// TIA Portal V20 export
// export: Created 2026-10-19T18:45:37.2686399Z, ExportSetting None, DisplayName Totally Integrated Automation Portal, DisplayVersion V20 Update 6, DisplayName TIA Portal Openness, DisplayVersion V20 Update 6, DisplayName TIA Portal Version Control Interface, DisplayVersion V20 Update 6, DisplayName SINAMICS Startdrive Advanced, DisplayVersion V20 SP1, DisplayName SINAMICS Startdrive G130, G150, S120, S150, SINAMICS MV, G220, S200, S210, DisplayVersion V20 SP1, DisplayName SINAMICS Startdrive G110M, G120, G120C, G120D, G120P, G115D, DisplayVersion V20 SP1, DisplayName STEP 7 Professional, DisplayVersion V20 Update 6, DisplayName STEP 7 Safety, DisplayVersion V20 Update 2, DisplayName WinCC Basic/Comfort/Advanced, DisplayVersion V20 Update 6, DisplayName WinCC Unified, DisplayVersion V20 Update 6
VAR_GLOBAL   // PLC tag table "IO_Remote_Panel_2"
   "KEY REMOTE/LOCAL L5 - CH1(2)" AT %I470.5 : Bool;
   "KEY REMOTE/LOCAL L2 - CH1(2)" AT %I461.7 : Bool;
   "VTD2 UPPER ULTIMATE CREEP" AT %I286.1 : Bool;
   "SAFETY_GATE_3_CH1(2)" AT %I461.2 : Bool;
   "STACK LIGHTS GREEN(2)" AT %Q174.3 : Bool;
   "C2112 VTD CIRCUIT BREAKER" AT %I285.0 : Bool;
   "STO VTD - CH1(2)" AT %Q446.2 : Bool;
   "STACK LIGHTS RED(2)" AT %Q174.1 : Bool;
   "LIGHT GUARDS 2 - CH2(2)" AT %I453.2 : Bool;
   "VTU HOIST BRAKE SAFETY ENABLE EDM FEEDBACK(2)" AT %I452.0 : Bool;
   "Chain Slack 3 - CH1(2)" AT %I356.6 : Bool;
   "KEY REMOTE/LOCAL L3 - CH1(2)" AT %I470.1 : Bool;
   "KEY REMOTE/LOCAL L6 - CH1(2)" AT %I470.7 : Bool;
   "BRAKE SUPPLY SAFETY CONTACTOR 1(2)" AT %Q446.0 : Bool;
   "KEY REMOTE/LOCAL L1 - CH2(2)" AT %I462.5 : Bool;
   "E-STOP L1 - CH2(2)" AT %I462.4 : Bool;
   "E-STOP L1 - CH1(2)" AT %I461.4 : Bool;
   "VTD2 PUSH TO EXIT VTD ZONE" AT %I286.6 : Bool;
   "E-STOP (CABINET) - CH1(2)" AT %I356.0 : Bool;
   "E-STOP L6 - CH2(2)" AT %I471.6 : Bool;
   "C2109, C2110, C2111 CVTD CIRCUIT BREAKER" AT %I285.3 : Bool;
   "E-STOP L2 - CH2(2)" AT %I462.6 : Bool;
   "SAFETY_GATE_1_CH2(2)" AT %I462.0 : Bool;
   "CABINET COOLING FAN CIRCUIT BREAKER FEEDBACK(2)" AT %I285.4 : Bool;
   "KEY REMOTE/LOCAL L6 - CH2(2)" AT %I471.7 : Bool;
   "STO VTD - CH2(2)" AT %Q446.3 : Bool;
   "KEY REMOTE/LOCAL L1 - CH1(2)" AT %I461.5 : Bool;
   "SAFETY_GATE_1_CH1(2)" AT %I461.0 : Bool;
   "KEY REMOTE/LOCAL L3 - CH2(2)" AT %I471.1 : Bool;
   "VTD2 UPPER ULTIMATE SLOWDOWN" AT %I286.0 : Bool;
   "VTD2 LOWER ULTIMATE SLOWDOWN" AT %I286.4 : Bool;
   "KEY REMOTE/LOCAL L4 - CH2(2)" AT %I471.3 : Bool;
   "E-STOP L6 - CH1(2)" AT %I470.6 : Bool;
   "KEY REMOTE/LOCAL L4 - CH1(2)" AT %I470.3 : Bool;
   "E-STOP L5 - CH1(2)" AT %I470.4 : Bool;
   "E-STOP L3 - CH2(2)" AT %I471.0 : Bool;
   "KEY REMOTE/LOCAL L5 - CH2(2)" AT %I471.5 : Bool;
   "BRAKE SUPPLY SAFETY CONTACTOR 2(2)" AT %Q446.1 : Bool;
   "SAFETY_GATE_4_CH1(2)" AT %I461.3 : Bool;
   "Chain Slack 3 - CH2(2)" AT %I357.6 : Bool;
   "STACK LIGHTS ORANGE(2)" AT %Q174.2 : Bool;
   "Chain Slack 2 - CH2(2)" AT %I357.5 : Bool;
   "C2105, C2106, C2107, C2108 CIRCUIT BREAKER" AT %I285.2 : Bool;
   "LIGHT GUARD 2 - CH1(2)" AT %I452.2 : Bool;
   "Chain Slack 2 - CH1(2)" AT %I356.5 : Bool;
   "KEY REMOTE/LOCAL L2 - CH2(2)" AT %I462.7 : Bool;
   "VTD2 PUSH TO ENTER VTD ZONE" AT %I286.5 : Bool;
   "CABINET 24V PSU CIRCUIT BREAKER FEEDBACK(2)" AT %I285.5 : Bool;
   "CABINET 24V PSU CIRCUIT BREAKER FEEDBACK_1(2)" AT %I285.6 : Bool;
   "Chain Slack 1 - CH1(2)" AT %I356.4 : Bool;
   "SAFETY_GATE_3_CH2(2)" AT %I462.2 : Bool;
   "RESET (CABINET)(2)" AT %I356.1 : Bool;
   "E-STOP L3 - CH1(2)" AT %I470.0 : Bool;
   "RESET LAMP(2)" AT %Q174.0 : Bool;   // TESTED
   "SAFETY_GATE_2_CH1(2)" AT %I461.1 : Bool;
   "E-STOP L5 - CH2(2)" AT %I471.4 : Bool;
   "VTD2 UPPER LIMIT" AT %I286.3 : Bool;
   "LIGHT GUARDS 1 - CH2(2)" AT %I453.1 : Bool;
   "Chain Slack 1 - CH2(2)" AT %I357.4 : Bool;
   "LIGHT GUARD 1 - CH1(2)" AT %I452.1 : Bool;
   "E-STOP L2 - CH1(2)" AT %I461.6 : Bool;
   "E-STOP L4 - CH2(2)" AT %I471.2 : Bool;
   "VTD2 LOWER LIMIT" AT %I286.2 : Bool;
   "SAFETY_GATE_4_CH2(2)" AT %I462.3 : Bool;
   "C2101, C2102, C2103, C2104 CIRCUIT BREAKER" AT %I285.1 : Bool;
   "E-STOP L4 - CH1(2)" AT %I470.2 : Bool;
   "E-STOP (CABINET) - CH2(2)" AT %I357.0 : Bool;
   "SAFETY_GATE_2_CH2(2)" AT %I462.1 : Bool;
   "Chain Slack 4 - CH2(2)" AT %I357.7 : Bool;
   "Chain Slack 4 - CH1(2)" AT %I356.7 : Bool;
   "RESET 2 PLC HMI" AT %Q174.5 : Bool;
   "PLC_HMI - HMI 2 Estop" AT %I357.2 : Bool;
   "PLC_HMI - HMI 1 Estop" AT %I356.2 : Bool;
   "PLC_HMI - Profinet_Error_HMI 1" AT %I356.3 : Bool;
   "PLC_HMI - Profinet_Error_HMI 2" AT %I357.3 : Bool;
   "RESET 1 PLC HMI" AT %Q174.4 : Bool;
END_VAR
